(* IEC 61131-3 sources: trust-platform/editors/vscode/src/test/fixtures/control-engineering/live-simulation-project/src, 1 file *)

(* ---- main.st ---- *)
USING Control;

PROGRAM Main
VAR
    Controller : Control.PID;
    Parameters : Control.PIDParameters;
    InitialState : Control.PIDInitialState;
    Input : Control.PIDInput;
    Initialized : BOOL := FALSE;
    AutoMode : BOOL := TRUE;
    Setpoint : LREAL := 20.0;
    ProcessValue : LREAL := 20.0;
    ManipulatedValue : LREAL := 13.3333333333;
    OptionalFeedback : LREAL := 0.0;
END_VAR

Parameters.ProportionalGain := LREAL#1.0;
Parameters.IntegralGain := LREAL#0.2;
Parameters.DerivativeGain := LREAL#0.0;
Parameters.ProportionalSetpointWeight := LREAL#1.0;
Parameters.DerivativeSetpointWeight := LREAL#0.0;
Parameters.Bias := LREAL#13.3333333333;
Parameters.OutputMinimum := LREAL#0.0;
Parameters.OutputMaximum := LREAL#100.0;
Parameters.RateMinimum := LREAL#-25.0;
Parameters.RateMaximum := LREAL#25.0;
Parameters.TrackingTime := LREAL#1.0;
Parameters.AntiWindup := PIDAntiWindup#Combined;

IF NOT Initialized THEN
    (* Configure once so an explicitly reviewed online parameter update is not
       overwritten by the startup constants on the following scan. *)
    Controller.Configure(Parameters := Parameters);
    InitialState.Setpoint := Setpoint;
    InitialState.ProcessValue := ProcessValue;
    InitialState.NominalOutput := ManipulatedValue;
    InitialState.SaturatedOutput := ManipulatedValue;
    Controller.Initialize(State := InitialState);
    Initialized := TRUE;
END_IF;

Input.Setpoint := Setpoint;
Input.ProcessValue := ProcessValue;
Input.Mode := PIDMode#Auto;
Input.CycleTime := LREAL#0.1;
ManipulatedValue := Controller.Update(Input := Input);
END_PROGRAM

CONFIGURATION Config
RESOURCE Res ON PLC
    TASK MainTask(INTERVAL := T#100ms, PRIORITY := 1);
    PROGRAM P1 WITH MainTask : Main;
END_RESOURCE
VAR_CONFIG
    P1.AutoMode AT %MX8.0 : BOOL;
    P1.Setpoint AT %ML0 : LREAL;
    P1.ManipulatedValue AT %QL0 : LREAL;
    P1.ProcessValue AT %IL0 : LREAL;
    P1.OptionalFeedback AT %IL8 : LREAL;
END_VAR
END_CONFIGURATION
